// TIA Portal V21 export
FUNCTION "FC_AnaOutputPath" : Void   // FC11, SCL
TITLE = Analyzer: output not written on every path
{ S7_Optimized_Access := 'TRUE' }
// Rule C26d: Result is not written when Select is FALSE
// stored: SetENOAutomatically false
   VAR_INPUT
      Select : Bool;   // Select the value
      Value : Int;   // Value
   END_VAR
   VAR_OUTPUT
      Result : Int;   // Result
   END_VAR
BEGIN

       IF #Select THEN
           #Result := #Value;
       END_IF;
END_FUNCTION
